(* Schneider Machine Expert - Basic project native_modbus_bare_abort_read_i, file version 3.0.0.0 *)
(* ProjectInformations: Name=New project *)

HARDWARE
  Cpu 0: TM200CE40T
  EthernetConfiguration: NetworkName=M200, IpAllocationMode=FixedAddress, IpAddress=0.0.0.0, SubnetMask=0.0.0.0
  SerialLineConfiguration: Baud=Baud19200, Parity=ParityEven, DataBits=DataBits8, StopBits=StopBits1, PhysicalMedium=PhysicalMediumRs485, TransmissionMode=TransmissionModeModbusRtu, SlaveId=1, Addressing=MasterAddressing
  MastTask: UsePeriodScanMode=false, PeriodScan=100
  FastTask: Period=255
  CpuBehavior: StartingMode=StartAsPreviousState, AutoSaveRamOnEeprom=true, WatchdogPeriod=250

SYMBOLS  (address, symbol, comment, settings)
  %READ_VAR0   [Link(Value(FBComLinkParameterEnums=SerialLine1)), RemoteDeviceId(Value(int=1)), Timeout(Value(int=100)), ObjType(Value(FBComObjTypeParameterEnums=I)), FirstObj(Value(int=17)), Quantity(Value(int=17)), IndexData(Value(int=200))]

POU Generated C++ - EXPERIMENTAL
  (* SectionNumber=0 *)

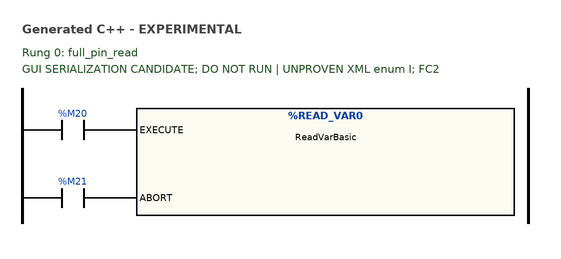

// Rung 0: full_pin_read
// GUI SERIALIZATION CANDIDATE; DO NOT RUN | UNPROVEN XML enum I; FC2
  BLK %READ_VAR0
  LD %M20
  EXECUTE
  LD %M21
  ABORT
  END_BLK
  // as ST:
  //   %READ_VAR0(EXECUTE := %M20, ABORT := %M21);
